// TIA Portal V19 export
FUNCTION_BLOCK "PUMP_FB1"   // FB5, FBD
{ S7_Optimized_Access := 'FALSE' }
// stored: SetENOAutomatically false
   VAR_INPUT
      "PUMP SELECTION" : Bool;
      TRIP : Bool;
      SIM : Bool;
      "AUTO START" : Bool;
   END_VAR
   VAR_OUTPUT
      OP_FBK_ERROR : Bool;
      CL_FBK_ERROR : Bool;
      AUTO_MODE : Bool;
      MANUAL_MODE : Bool;
      SEMI_AUTO_MODE : Bool;
      "START/STOPCMD" : Bool;
      STATUS : Int;
      FAULT : Bool;
   END_VAR
   VAR_IN_OUT
      "MANUAL SELECTION" : Bool;
      SEMI : Bool;
      "MANUAL START" : Bool;
      "FEEDBACK RUN" : Bool;
      TRIPPED : Bool;
      REMOTE : Bool;
      RESET : Bool;
      INTERLOCK : Bool;
      "WAITING TIME" : DInt;
   END_VAR
   VAR
      "TIMER" { S7_SetPoint := 'True'} : IEC_TIMER;
      MON_ERROR : Bool;
      INTERLOCK_ACTIVE : Bool;
      SIM_FBK_RUN : Bool;
   END_VAR
   // "TIMER".PT := T#10S;
   VAR_TEMP   // added for the SCL form of the ladder/FBD networks
      _w1 : Bool;
   END_VAR
BEGIN

REGION Network 1: MODE SELECTION
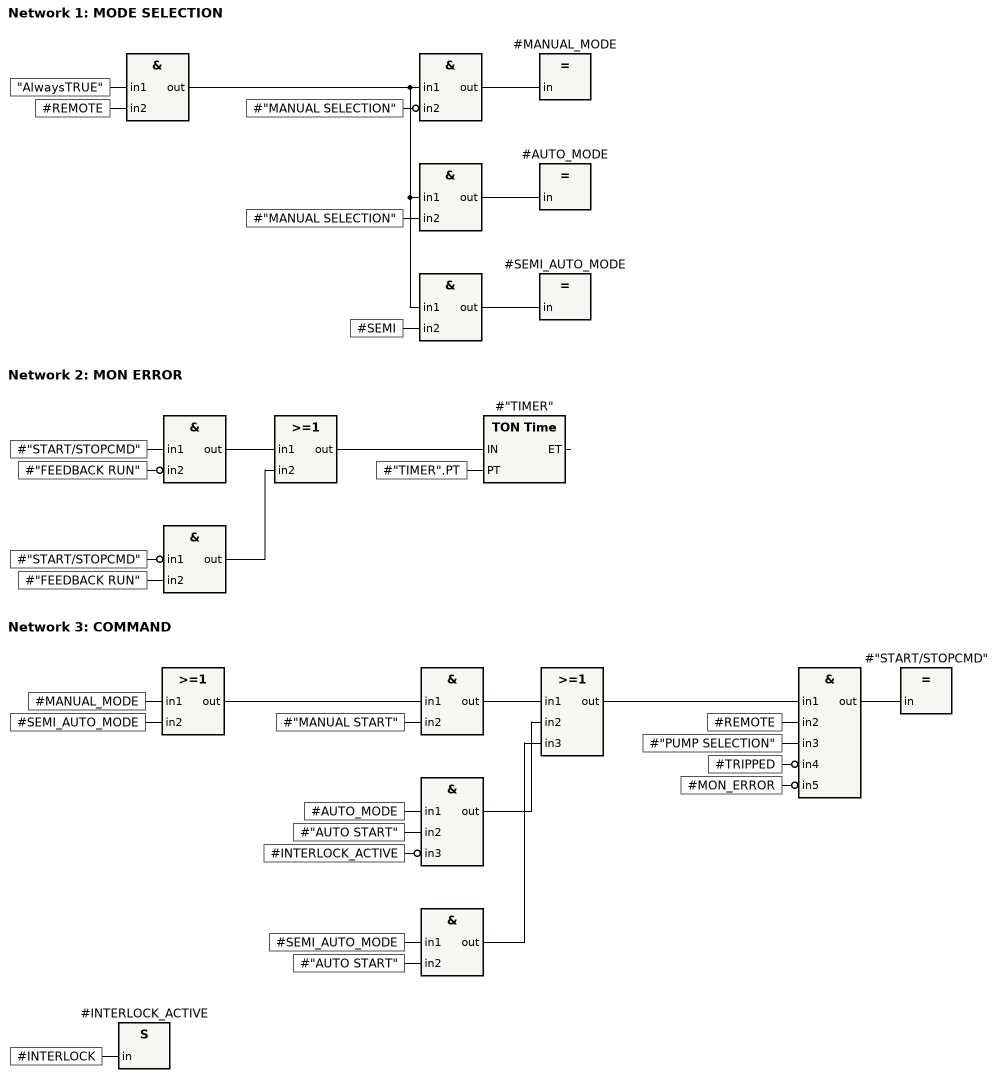
   #_w1 := "AlwaysTRUE" AND #REMOTE;
   #MANUAL_MODE := #_w1 AND NOT #"MANUAL SELECTION";
   #AUTO_MODE := #_w1 AND #"MANUAL SELECTION";
   #SEMI_AUTO_MODE := #_w1 AND #SEMI;
END_REGION

REGION Network 2: MON ERROR
   #"TIMER".TON(IN := (#"START/STOPCMD" AND NOT #"FEEDBACK RUN") OR (NOT #"START/STOPCMD" AND #"FEEDBACK RUN"),
                PT := #"TIMER".PT);
END_REGION

REGION Network 3: COMMAND
   #"START/STOPCMD" := (((#MANUAL_MODE OR #SEMI_AUTO_MODE) AND #"MANUAL START") OR (#AUTO_MODE AND #"AUTO START" AND NOT #INTERLOCK_ACTIVE) OR (#SEMI_AUTO_MODE AND #"AUTO START")) AND #REMOTE AND #"PUMP SELECTION" AND NOT #TRIPPED AND NOT #MON_ERROR;
   IF #INTERLOCK THEN #INTERLOCK_ACTIVE := TRUE; END_IF;
END_REGION

REGION Network 4: MON ERROR
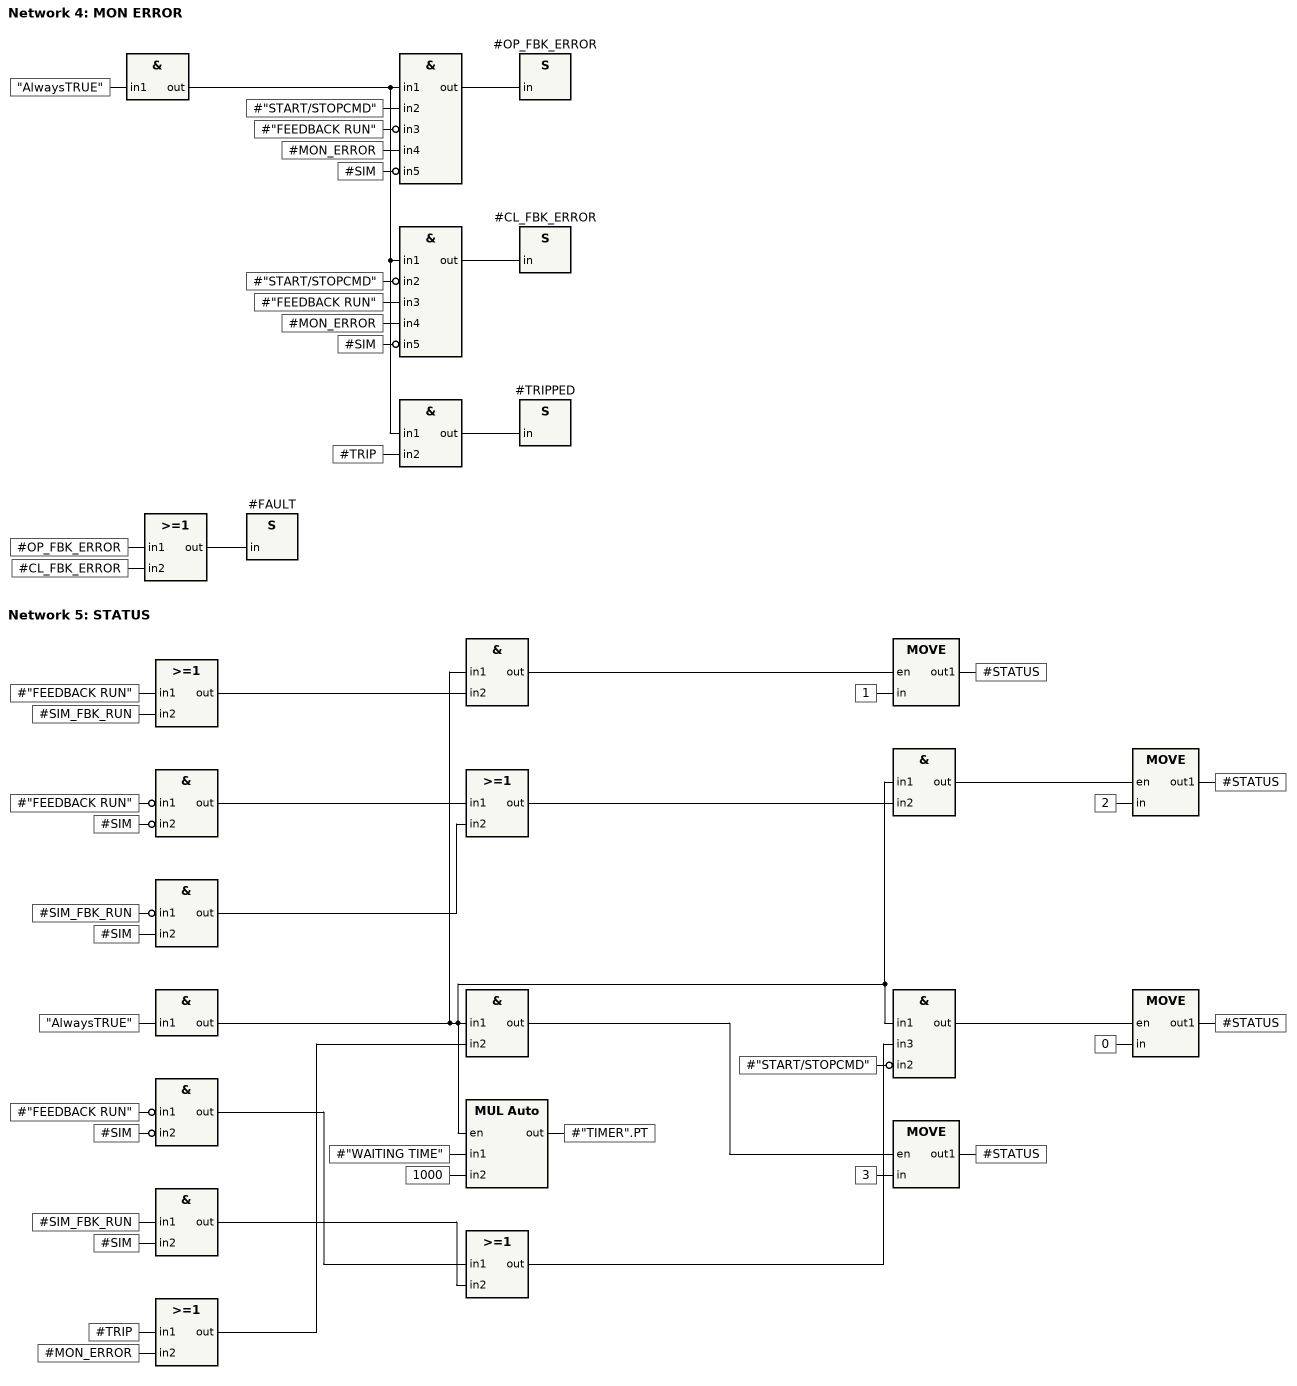
   IF "AlwaysTRUE" AND #"START/STOPCMD" AND NOT #"FEEDBACK RUN" AND #MON_ERROR AND NOT #SIM THEN
       #OP_FBK_ERROR := TRUE;
   END_IF;
   IF "AlwaysTRUE" AND NOT #"START/STOPCMD" AND #"FEEDBACK RUN" AND #MON_ERROR AND NOT #SIM THEN
       #CL_FBK_ERROR := TRUE;
   END_IF;
   IF "AlwaysTRUE" AND #TRIP THEN #TRIPPED := TRUE; END_IF;
   IF #OP_FBK_ERROR OR #CL_FBK_ERROR THEN #FAULT := TRUE; END_IF;
END_REGION

REGION Network 5: STATUS
   IF "AlwaysTRUE" AND (#"FEEDBACK RUN" OR #SIM_FBK_RUN) THEN #STATUS := 1; END_IF;
   IF "AlwaysTRUE" AND ((NOT #"FEEDBACK RUN" AND NOT #SIM) OR (NOT #SIM_FBK_RUN AND #SIM)) THEN
       #STATUS := 2;
   END_IF;
   IF "AlwaysTRUE" AND ((NOT #"FEEDBACK RUN" AND NOT #SIM) OR (#SIM_FBK_RUN AND #SIM)) AND NOT #"START/STOPCMD" THEN
       #STATUS := 0;
   END_IF;
   IF "AlwaysTRUE" AND (#TRIP OR #MON_ERROR) THEN #STATUS := 3; END_IF;
   IF "AlwaysTRUE" THEN #"TIMER".PT := #"WAITING TIME" * 1000; END_IF;
END_REGION

REGION Network 6: RESET
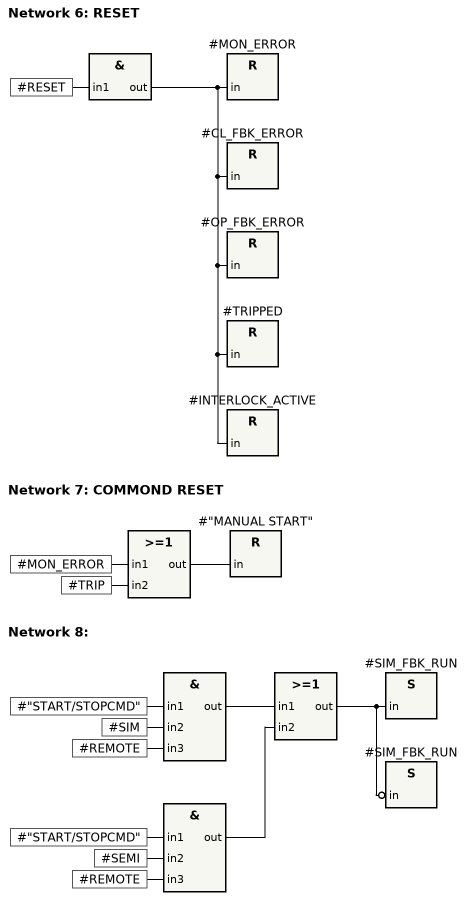
   IF #RESET THEN
       #MON_ERROR := FALSE;
       #CL_FBK_ERROR := FALSE;
       #OP_FBK_ERROR := FALSE;
       #TRIPPED := FALSE;
       #INTERLOCK_ACTIVE := FALSE;
   END_IF;
END_REGION

REGION Network 7: COMMOND RESET
   IF #MON_ERROR OR #TRIP THEN #"MANUAL START" := FALSE; END_IF;
END_REGION

REGION Network 8
   #_w1 := (#"START/STOPCMD" AND #SIM AND #REMOTE) OR (#"START/STOPCMD" AND #SEMI AND #REMOTE);
   IF #_w1 THEN #SIM_FBK_RUN := TRUE; END_IF;
   IF NOT #_w1 THEN #SIM_FBK_RUN := TRUE; END_IF;
END_REGION
END_FUNCTION_BLOCK
